Fanuc KAREL source: KA00090.KL

PROGRAM KA00090
%NOLOCKGROUP
VAR
  SRC: JOINTPOS
  DST: XYZWPR
BEGIN
  DST = SRC
END KA00090
